(* IEC 61131-3 sources: plc-vscode/tests/st/all/trust-platform/examples/OSCAT/tunnel_washer_chain/non-oop/src, 3 files *)

(* ---- Main.st ---- *)
FUNCTION_BLOCK ClassicWasherQuality
VAR
    LastHandlerIdValue : INT;
    RejectCounter : DwordCounter;
END_VAR

METHOD PUBLIC Initialize
RejectCounter.Initialize();
RejectCounter.Configure(StepSize := DWORD#1, MaxValue := DWORD#16#FFFFFFFF);
END_METHOD

METHOD PUBLIC Evaluate : INT
VAR_INPUT
    SoilLevel : REAL;
    Conductivity : REAL;
    RinseConductivity : REAL;
    OperatorAvailable : BOOL;
END_VAR
IF (SoilLevel > REAL#70.0) AND (Conductivity < REAL#3.0) THEN
    LastHandlerIdValue := INT#1;
ELSIF RinseConductivity > REAL#1.5 THEN
    LastHandlerIdValue := INT#2;
ELSIF OperatorAvailable THEN
    LastHandlerIdValue := INT#3;
ELSE
    LastHandlerIdValue := INT#4;
    RejectCounter.Update(Up := TRUE, Down := FALSE);
END_IF;
Evaluate := LastHandlerIdValue;
END_METHOD

PUBLIC PROPERTY RejectCount : DWORD
GET
    RejectCount := RejectCounter.Count;
END_GET
END_PROPERTY
END_FUNCTION_BLOCK

PROGRAM Main
VAR
    Washer : ClassicWasherQuality;
    Handler : INT;
END_VAR
Washer.Initialize();
Handler := Washer.Evaluate(SoilLevel := REAL#80.0, Conductivity := REAL#2.0, RinseConductivity := REAL#0.5, OperatorAvailable := FALSE);
END_PROGRAM

(* ---- Configuration.st ---- *)
CONFIGURATION TunnelWasherChainClassicConfiguration
RESOURCE Cpu0 ON PLC
    TASK MainTask (INTERVAL := T#100ms, PRIORITY := 1);
    PROGRAM Washer WITH MainTask : Main;
END_RESOURCE
END_CONFIGURATION

(* ---- Tests.st ---- *)
TEST_PROGRAM ClassicWasherFallsThroughToReject
VAR
    Washer : ClassicWasherQuality;
END_VAR

Washer.Initialize();
ASSERT_EQUAL(EXPECTED := INT#4, ACTUAL := Washer.Evaluate(SoilLevel := REAL#40.0, Conductivity := REAL#4.0, RinseConductivity := REAL#0.5, OperatorAvailable := FALSE));
ASSERT_EQUAL(EXPECTED := DWORD#1, ACTUAL := Washer.RejectCount);
END_TEST_PROGRAM
